Staubli VAL3: main.pgx

program main()
begin
  close(tCurrentTool)
  pPointRs.config.shoulder = lefty
  pPointRs2.config.shoulder = lefty
  mCurrentSpeed.tvel = 100.00
  mCurrentSpeed.blend = joint
  mCurrentSpeed.reach = 0.010
  mCurrentSpeed.leave = 0.010
  // Program PgProg start
  // Program generated by RoboDK v6.0.7 for Staubli TS20 FL 100 TC on XX/XX/XXXX 18:00:00
  // Using nominal kinematics.
  mCurrentSpeed.tvel = 250.000
  mCurrentSpeed.reach = 5.000
  mCurrentSpeed.leave = 5.000
  call MoveJoint(10.00000,-20.00000,50.00000,30.00000)
  call MoveLine(-607.850,543.849,363.215,136.262,30.757,-130.375)
  call MoveCirc(-602.951,596.788,316.595,136.262,30.757,-130.375,-663.517,575.988,286.611,136.262,30.757,-130.375)
  call MoveJoint(30.00000,25.00000,80.00000,-45.00000)
  mCurrentSpeed.tvel = 100.000
  call MoveLine(-650.861,503.437,361.399,136.262,30.757,-130.375)
  mCurrentSpeed.reach = 0.000
  mCurrentSpeed.leave = 0.000
  call MoveLine(-640.584,506.980,371.534,136.262,30.757,-130.375)
  delay(0.500)
  popUpMsg("Paused. Press OK to continue")
  popUpMsg("Hello from postgen")
  // a comment
  //call prog:SubProgram()
  CustomCode(42)
  ThreadProg
  Output[1]=true
  Valve=false
  Output[3]=2.5
  watch(Input[2]==true)
  watch(Input[4]==false,1500.0)
  call MoveJoint(10.00000,-20.00000,50.00000,30.00000)
  call MoveJoint(20.00000,-15.00000,55.00000,35.00000)
  call MoveLine(-353.026,-90.135,331.702,164.619,39.324,-168.579)

  waitEndMove()
  // Program PgProg end

end
